(* CODESYS project P_Settings.xml

Project tree, tasks and I/O mapping:
*)

// P_Settings
PROPERTY P_Settings : REFERENCE TO ST_AlarmSettings
END_PROPERTY
